(* IEC 61131-3 sources: RootPLC/conformance/cases/types, 56 files *)

(* ---- err_struct_recursive.st ---- *)
(* spec: [types.derived.struct]
   expect: error RP0107 *)
TYPE N : STRUCT child : N; END_STRUCT; END_TYPE

(* ---- err_subrange_bounds.st ---- *)
(* spec: [types.derived.subrange]
   expect: error RP0108 *)
TYPE Bad : INT (10..0); END_TYPE

(* ---- ok_call_through_reference.st ---- *)
(* spec: [types.reference.alias] [pous.call.callee]
   expect: warning RP0118
   run: PRG_Main cycles=2
   assert: c.n = 4 *)
FUNCTION_BLOCK FB_Count
VAR_OUTPUT
    n : INT;
END_VAR
n := n + 1;
END_FUNCTION_BLOCK

PROGRAM PRG_Main
VAR
    c : FB_Count;
    r : REFERENCE TO FB_Count;
END_VAR
r REF= c;
r();          (* calls c through the reference *)
c();
END_PROGRAM

(* ---- err_array_bound_not_constant.st ---- *)
(* spec: [variables.constant-names]
   expect: error RP0108 *)
PROGRAM PRG_Main
VAR
    n : INT := 4;
    buffer : ARRAY[0..n] OF INT;
END_VAR
END_PROGRAM

(* ---- err_array_bounds.st ---- *)
(* spec: [types.derived.array]
   expect: error RP0108 *)
PROGRAM PRG_Main
VAR
    a : ARRAY[5..1] OF INT;
END_VAR

END_PROGRAM

(* ---- err_array_const_index.st ---- *)
(* spec: [types.derived.array]
   expect: error RP0109 *)
PROGRAM PRG_Main
VAR
    a : ARRAY[0..2] OF INT;
END_VAR
a[3] := 1;
END_PROGRAM

(* ---- err_const_overflow.st ---- *)
(* spec: [types.int.overflow]
   expect: error RP0101 *)
PROGRAM PRG_Main
VAR
    x : LINT := 9223372036854775807 + 1;
END_VAR

END_PROGRAM

(* ---- err_dint_to_real.st ---- *)
(* spec: [types.conversion.implicit]
   expect: error RP0103 *)
PROGRAM PRG_Main
VAR
    r : REAL;
    d : DINT;
END_VAR
r := d;
END_PROGRAM

(* ---- err_div_const_zero.st ---- *)
(* spec: [types.int.division]
   expect: error RP0101 *)
PROGRAM PRG_Main
VAR
    x : INT;
END_VAR
x := 5 / 0;
END_PROGRAM

(* ---- err_enum_ambiguous.st ---- *)
(* spec: [types.derived.enum]
   expect: error RP0106 *)
TYPE Mode : (Off, Manual, Auto); END_TYPE

TYPE Valve : (Closed, Auto); END_TYPE

PROGRAM PRG_Main
VAR
    i : INT;
END_VAR
i := TO_INT(Auto);   (* no expected enumeration: Mode#Auto or Valve#Auto? *)
END_PROGRAM

(* ---- err_enum_strict_assign.st ---- *)
(* spec: [types.derived.enum.integer]
   expect: error RP0103 *)
{attribute 'qualified_only'}
{attribute 'strict'}
TYPE StrictMode : (Idle, Busy);
END_TYPE

PROGRAM PRG_Main
VAR
    s : StrictMode;
    i : INT := 1;
END_VAR
s := i;       (* an integer variable cannot be stored in a strict enumeration *)
i := s + 1;   (* no arithmetic on a strict enumeration *)
END_PROGRAM

(* ---- err_generic_decl.st ---- *)
(* spec: [types.generic]
   expect: error RP0104 *)
PROGRAM PRG_Main
VAR
    x : ANY_INT;
END_VAR

END_PROGRAM

(* ---- err_implicit_narrowing.st ---- *)
(* spec: [types.conversion.implicit]
   expect: error RP0103 *)
PROGRAM PRG_Main
VAR
    si : SINT;
    i : INT := 1;
END_VAR
si := i;
END_PROGRAM

(* ---- err_index_non_array.st ---- *)
(* spec: [types.derived.array]
   expect: error RP0103 *)
(* Only arrays (and, as vendor forms, strings and references) can be
   indexed. *)
PROGRAM PRG_Main
VAR
    x : INT;
    y : INT;
END_VAR
y := x[0];
END_PROGRAM

(* ---- err_int_to_bool.st ---- *)
(* spec: [types.conversion.implicit]
   expect: error RP0103 *)
PROGRAM PRG_Main
VAR
    b : BOOL;
    i : INT := 1;
END_VAR
b := i;
END_PROGRAM

(* ---- err_literal_range.st ---- *)
(* spec: [types.literal.range]
   expect: error RP0102 *)
PROGRAM PRG_Main
VAR
    x : SINT := 200;
END_VAR

END_PROGRAM

(* ---- err_string_len_zero.st ---- *)
(* spec: [types.derived.string]
   expect: error RP0108 *)
PROGRAM PRG_Main
VAR
    s : STRING[0];
END_VAR

END_PROGRAM

(* ---- err_struct_name_equivalence.st ---- *)
(* spec: [types.equivalence] [types.derived.struct]
   expect: error RP0103 *)
TYPE A : STRUCT v : INT; END_STRUCT; END_TYPE
TYPE B : STRUCT v : INT; END_STRUCT; END_TYPE

PROGRAM PRG_Main
VAR
    a : A;
    b : B;
END_VAR
a := b;
END_PROGRAM

(* ---- err_subrange_const.st ---- *)
(* spec: [types.derived.subrange]
   expect: error RP0105 *)
TYPE Percent : INT (0..100); END_TYPE

PROGRAM PRG_Main
VAR
    p : Percent := 150;
END_VAR

END_PROGRAM

(* ---- err_unknown_type.st ---- *)
(* spec: [types.derived.alias]
   expect: error RP0111 *)
PROGRAM PRG_Main
VAR
    x : NoSuchType;
END_VAR

END_PROGRAM

(* ---- ok_alias.st ---- *)
(* spec: [types.derived.alias] [types.equivalence]
   expect: ok
   run: PRG_Main cycles=1
   assert: i = 10
   assert: s = 11 *)
TYPE Speed : INT := 10; END_TYPE

PROGRAM PRG_Main
VAR
    s : Speed;
    i : INT;
END_VAR
i := s;
s := i + 1;
END_PROGRAM

(* ---- ok_array.st ---- *)
(* spec: [types.derived.array]
   expect: ok
   run: PRG_Main cycles=1
   assert: a[2] = 7
   assert: a[0] = 0
   assert: m[2, 2] = TRUE *)
PROGRAM PRG_Main
VAR
    a : ARRAY[0..2] OF INT;
    m : ARRAY[1..2, 1..2] OF BOOL;
END_VAR
a[2] := 7;
m[2, 2] := TRUE;
END_PROGRAM

(* ---- ok_conv_to_string.st ---- *)
(* spec: [types.conversion.explicit]
   expect: ok
   run: PRG_Main cycles=1
   assert: a = '42'
   assert: b = '255'
   assert: c = 'T#1s500ms'
   assert: d = 'A'
   assert: e = 'TRUE'
   assert: f = '-7' *)
PROGRAM PRG_Main
VAR
    a, b, c, d, e, f : STRING;
    ch : CHAR := CHAR#'A';
END_VAR
a := INT_TO_STRING(42);
b := WORD_TO_STRING(16#FF);
c := TIME_TO_STRING(T#1500MS);
d := CHAR_TO_STRING(ch);
e := BOOL_TO_STRING(TRUE);
f := DINT_TO_STRING(-7);
END_PROGRAM

(* ---- ok_datetime_to_string.st ---- *)
(* spec: [types.conversion.explicit]
   expect: ok
   run: PRG_Main cycles=1
   assert: sDt = 'DT#2017-04-04-12:42:42'
   assert: sD = 'D#1999-12-31'
   assert: sTod = 'TOD#08:05:03.25'
   assert: sB = 'TRUE'
   assert: sI = '-42' *)
PROGRAM PRG_Main
VAR
    sDt, sD, sTod, sB, sI : STRING;
END_VAR
sDt := DT_TO_STRING(DT#2017-04-04-12:42:42);
sD := DATE_TO_STRING(D#1999-12-31);
sTod := TOD_TO_STRING(TOD#08:05:03.25);
sB := BOOL_TO_STRING(TRUE);
sI := INT_TO_STRING(-42);
END_PROGRAM

(* ---- ok_default_init.st ---- *)
(* spec: [types.elementary] [types.default-init]
   expect: ok
   run: PRG_Main cycles=1
   assert: b = FALSE
   assert: i = 0
   assert: u = 0
   assert: r = 0.0
   assert: w = 0
   assert: t = T#0s
   assert: lt = LT#0s
   assert: d = D#1970-01-01
   assert: s = ''
   assert: ws = "" *)
PROGRAM PRG_Main
VAR
    b : BOOL;
    i : INT;
    u : ULINT;
    r : LREAL;
    w : WORD;
    t : TIME;
    lt : LTIME;
    d : DATE;
    s : STRING;
    ws : WSTRING;
END_VAR

END_PROGRAM

(* ---- ok_enum.st ---- *)
(* spec: [types.derived.enum]
   expect: ok
   run: PRG_Main cycles=1
   assert: first = Mode#Off
   assert: m = Mode#Auto
   assert: i = 2 *)
TYPE Mode : (Off, Manual, Auto); END_TYPE

PROGRAM PRG_Main
VAR
    m : Mode;
    first : Mode;
    i : INT;
END_VAR
first := m;
m := Manual;
m := Mode#Auto;
i := TO_INT(m);
END_PROGRAM

(* ---- ok_enum_value_by_context.st ---- *)
(* spec: [types.derived.enum]
   expect: ok
   run: PRG_Main cycles=1
   assert: n = 2
   assert: hit = TRUE
   assert: m = Motor#RUN
   assert: d = Door#OPEN *)
TYPE Motor : (IDLE, RUN, FAULT);
END_TYPE

TYPE Door : (IDLE, OPEN, CLOSED);
END_TYPE

FUNCTION F_Open : BOOL
VAR_INPUT
    d : Door;
END_VAR
F_Open := d = OPEN;
END_FUNCTION

PROGRAM PRG_Main
VAR
    m : Motor := IDLE;     (* initial value: Motor#IDLE *)
    d : Door;
    n : INT;
    hit : BOOL;
END_VAR
IF m = IDLE THEN           (* comparison: the other operand decides *)
    m := RUN;              (* assignment: the target decides *)
END_IF;
CASE m OF
    IDLE: n := 1;          (* CASE label: the selector decides *)
    RUN: n := 2;
END_CASE;
d := OPEN;
hit := F_Open(IDLE) = FALSE AND F_Open(d);   (* parameter decides *)
END_PROGRAM

(* ---- ok_explicit_conversion.st ---- *)
(* spec: [types.conversion.explicit]
   expect: ok
   run: PRG_Main cycles=1
   assert: a = 44
   assert: b = 3
   assert: c = -3
   assert: d = 127
   assert: e = -3 *)
PROGRAM PRG_Main
VAR
    a : SINT;
    b : INT;
    c : INT;
    d : SINT;
    e : INT;
END_VAR
a := INT_TO_SINT(300);
b := REAL_TO_INT(2.5);
c := REAL_TO_INT(-2.5);
d := LREAL_TO_SINT(1000.0);
e := TO_INT(SINT#-3);
END_PROGRAM

(* ---- ok_implicit_widening.st ---- *)
(* spec: [types.conversion.implicit]
   expect: ok
   run: PRG_Main cycles=1
   assert: i = -5
   assert: d = -5.0
   assert: w = 15 *)
PROGRAM PRG_Main
VAR
    s : SINT := -5;
    i : INT;
    d : LREAL;
    b : BYTE := 16#0F;
    w : WORD;
END_VAR
i := s;
d := i;
w := b;
END_PROGRAM

(* ---- ok_int_division.st ---- *)
(* spec: [types.int.division]
   expect: ok
   run: PRG_Main cycles=1
   assert: a = -3
   assert: b = -1
   assert: c = 1 *)
PROGRAM PRG_Main
VAR
    a : INT;
    b : INT;
    c : INT;
END_VAR
a := -7 / 2;
b := -7 MOD 2;
c := 7 MOD -2;
END_PROGRAM

(* ---- ok_int_wrap.st ---- *)
(* spec: [types.int.overflow]
   expect: ok
   run: PRG_Main cycles=1
   assert: x = -128
   assert: u = 255 *)
PROGRAM PRG_Main
VAR
    x : SINT := 127;
    u : USINT := 0;
END_VAR
x := x + 1;
u := u - 1;
END_PROGRAM

(* ---- ok_real_no_fault.st ---- *)
(* spec: [types.real]
   expect: ok
   run: PRG_Main cycles=1
   assert: big = TRUE *)
PROGRAM PRG_Main
VAR
    r : LREAL := 1.0;
    big : BOOL;
END_VAR
r := r / 0.0;
big := r > 1.0E308;
END_PROGRAM

(* ---- ok_reference.st ---- *)
(* spec: [types.reference]
   expect: ok
   run: PRG_Main cycles=1
   assert: x = 9 *)
PROGRAM PRG_Main
VAR
    x : INT := 5;
    r : REF_TO INT;
END_VAR
r := REF(x);
r^ := 9;
END_PROGRAM

(* ---- ok_string_truncate.st ---- *)
(* spec: [types.derived.string]
   expect: ok
   run: PRG_Main cycles=1
   assert: s = 'abcde' *)
PROGRAM PRG_Main
VAR
    s : STRING[5];
    t : STRING := 'abcdefgh';
END_VAR
s := t;
END_PROGRAM

(* ---- ok_struct.st ---- *)
(* spec: [types.derived.struct] [types.reference]
   expect: ok
   run: PRG_Main cycles=1
   assert: p.x = 1
   assert: p.y = 0
   assert: n.next = NULL *)
TYPE Point : STRUCT x : INT := 1; y : INT; END_STRUCT; END_TYPE
TYPE Node : STRUCT next : REF_TO Node; v : INT; END_STRUCT; END_TYPE

PROGRAM PRG_Main
VAR
    p : Point;
    n : Node;
END_VAR

END_PROGRAM

(* ---- ok_subrange.st ---- *)
(* spec: [types.derived.subrange]
   expect: ok
   run: PRG_Main cycles=1
   assert: first = 0
   assert: p = 50 *)
TYPE Percent : INT (0..100); END_TYPE

PROGRAM PRG_Main
VAR
    p : Percent;
    first : INT;
END_VAR
first := p;
p := 50;
END_PROGRAM

(* ---- ok_time_arithmetic.st ---- *)
(* spec: [types.time.arith]
   expect: ok
   run: PRG_Main cycles=1
   assert: t1 = TOD#08:30:00
   assert: t2 = TOD#23:30:00
   assert: d1 = DT#2026-11-04-12:01:30
   assert: d2 = DT#2026-11-04-11:59:00
   assert: dur1 = T#90000ms
   assert: dur2 = T#86400000ms
   assert: dur3 = T#3600000ms
   assert: lt = LTOD#00:00:01 *)
PROGRAM PRG_Main
VAR
    t1, t2 : TOD;
    d1, d2 : DT;
    dur1, dur2, dur3 : TIME;
    lt : LTOD;
END_VAR
t1 := TOD#08:00:00 + T#30M;
t2 := TOD#00:30:00 - T#1H;                        (* wraps around midnight *)
d1 := DT#2026-11-04-12:00:00 + T#1M30S500MS;      (* whole seconds *)
d2 := DT#2026-11-04-12:00:00 - T#1M;
dur1 := DT#2026-11-04-12:01:30 - DT#2026-11-04-12:00:00;
dur2 := D#2026-11-05 - D#2026-11-04;
dur3 := TOD#13:00:00 - TOD#12:00:00;
lt := LTOD#23:59:59 + LT#2S;
END_PROGRAM

(* ---- ok_time_conversions.st ---- *)
(* spec: [types.conversion.explicit] [types.conversion.implicit]
   expect: ok
   run: PRG_Main cycles=1
   assert: toL = LT#3ms
   assert: toT = T#1ms
   assert: viaTo = T#10ms
   assert: widened = LT#250ms
   assert: initL = LT#2s
   assert: atLdt = LDT#2026-01-01-10:00:00
   assert: atDt = DT#2026-01-01-10:00:00
   assert: atLtod = LTOD#12:30:00
   assert: gt = TRUE
   assert: eq = TRUE
   assert: later = TRUE
   assert: biggest = LT#2ms
   assert: ns = 1000000 *)
PROGRAM PRG_Main
VAR
    t : TIME := T#250ms;
    initL : LTIME := T#2s;
    toL, widened, biggest : LTIME;
    toT, viaTo : TIME;
    atLdt : LDT;
    atDt : DT;
    atLtod : LTOD;
    gt, eq, later : BOOL;
    ns : ULINT;
END_VAR
toL := TIME_TO_LTIME(T#3ms);
toT := LTIME_TO_TIME(LT#1500us);
viaTo := TO_TIME(TO_LTIME(UDINT#100000 * 100));
widened := t;
atLdt := DT#2026-01-01-10:00:00;
atDt := TO_DT(LDT#2026-01-01-10:00:00);
atLtod := TOD#12:30:00;
gt := T#2ms > LT#1ms;
eq := T#2ms = LT#2ms;
later := DT#2026-01-01-00:00:00 > LDT#2025-01-01-00:00:00;
biggest := MAX(T#2ms, LT#1ms);
ns := LTIME_TO_ULINT(T#1ms);
END_PROGRAM

(* ---- ok_to_string_forms.st ---- *)
(* spec: [types.conversion.explicit]
   expect: ok
   run: PRG_Main cycles=1
   assert: r1 = '0.1'
   assert: r2 = '-3.402823E38'
   assert: r3 = '1.0'
   assert: l1 = '123456789.0'
   assert: l2 = '1E-7'
   assert: t1 = 'T#49d17h2m47s295ms'
   assert: t2 = 'T#1s500ms'
   assert: t3 = 'T#0ms'
   assert: t4 = 'LT#1ms500us' *)
PROGRAM PRG_Main
VAR
    r1, r2, r3, l1, l2 : STRING;
    t1, t2, t3, t4 : STRING;
END_VAR
r1 := REAL_TO_STRING(REAL#0.1);
r2 := REAL_TO_STRING(REAL#-3.402823E38);
r3 := REAL_TO_STRING(REAL#1.0);
l1 := LREAL_TO_STRING(123456789.0);
l2 := LREAL_TO_STRING(1.0E-7);
t1 := TIME_TO_STRING(T#49d17h2m47s295ms);
t2 := TIME_TO_STRING(T#1500ms);
t3 := TIME_TO_STRING(T#0ms);
t4 := LTIME_TO_STRING(LTIME#1500us);
END_PROGRAM

(* ---- ok_untyped_literal.st ---- *)
(* spec: [types.literal.untyped]
   expect: ok
   run: PRG_Main cycles=1
   assert: u = 255
   assert: r = 3.0 *)
PROGRAM PRG_Main
VAR
    u : USINT := 255;
    r : REAL := 3;
END_VAR

END_PROGRAM

(* ---- warn_adr.st ---- *)
(* spec: [types.reference]
   expect: warning RP0117
   run: PRG_Main cycles=1
   assert: v = 9 *)
PROGRAM PRG_Main
VAR
    x : INT := 4;
    r : REF_TO INT;
    v : INT;
END_VAR
r := ADR(x);
r^ := 9;
v := x;
END_PROGRAM

(* ---- warn_array_bound_enum.st ---- *)
(* spec: [variables.constant-names] [scope.vendor-forms]
   expect: warning RP0135
   run: PRG_Main cycles=1
   assert: lo = 1
   assert: hi = 3
   assert: n = 3 *)
TYPE ST_Lanes :
STRUCT
    speed : ARRAY[E_Lane.Nr1..E_Lane.Nr3] OF INT;
END_STRUCT;
END_TYPE

TYPE E_Lane : (Nr1 := 1, Nr2, Nr3); END_TYPE

PROGRAM PRG_Main
VAR
    lanes : ARRAY[E_Lane.Nr1..E_Lane.Nr3] OF INT;
    lanes2 : ST_Lanes;
    lo, hi, n : DINT;
END_VAR
lo := LOWER_BOUND(lanes, 1);
hi := UPPER_BOUND(lanes, 1);
n := UPPER_BOUND(lanes2.speed, 1);
END_PROGRAM

(* ---- warn_enum_as_integer.st ---- *)
(* spec: [types.derived.enum.integer]
   expect: warning RP0129
   run: PRG_Main cycles=1
   assert: n = 2
   assert: plus = 3
   assert: next = Mode#Auto
   assert: same = TRUE
   assert: k = 1
   assert: fromInt = Mode#Manual
   assert: big = TRUE *)
TYPE Mode : (Off, Manual, Auto);
END_TYPE

TYPE Level : (Low, Mid, High);
END_TYPE

{attribute 'strict'}
TYPE StrictMode : (Idle, Busy);
END_TYPE

PROGRAM PRG_Main
VAR
    m : Mode := Mode#Auto;
    n : INT;
    plus : INT;
    next : Mode;
    same : BOOL;
    k : INT;
    fromInt : Mode;
    i : INT := 1;
    s : StrictMode;
    big : BOOL;
END_VAR
n := m;                           (* value as integer *)
plus := Mode#Auto + 1;            (* arithmetic on a non-strict enumeration *)
next := Mode#Manual + 1;          (* integer stored in a non-strict enumeration *)
same := Mode#Auto = Level#High;   (* compared as integers *)
s := StrictMode#Busy;
k := s;                           (* a strict value still reads as an integer *)
big := s > 0;
fromInt := i;
END_PROGRAM

(* ---- warn_enum_base_type_after.st ---- *)
(* spec: [types.derived.enum]
   expect: warning RP0115
   run: PRG_Main cycles=1
   assert: n = 10 *)
TYPE E_Mode : (Off := 0, Manual := 5, Auto := 10) UINT; END_TYPE

PROGRAM PRG_Main
VAR
    m : E_Mode := E_Mode#Auto;
    n : INT;
END_VAR
n := TO_INT(m);
END_PROGRAM

(* ---- warn_enum_dot_value.st ---- *)
(* spec: [types.derived.enum]
   expect: warning RP0122
   run: PRG_Main cycles=1
   assert: n = 10
   assert: same = TRUE
   assert: k = 1 *)
TYPE E_Mode : (Off := 0, Manual := 5, Auto := 10); END_TYPE

NAMESPACE Plant
TYPE E_Valve : (Closed, Open); END_TYPE
END_NAMESPACE

PROGRAM PRG_Main
VAR
    m : E_Mode := E_Mode.Auto;
    v : Plant.E_Valve;
    n, k : INT;
    same : BOOL;
END_VAR
n := TO_INT(m);
same := m = E_Mode#Auto;
v := Plant.E_Valve.Open;
k := TO_INT(v);
END_PROGRAM

(* ---- warn_enum_to_int.st ---- *)
(* spec: [types.derived.enum] [types.derived.enum.integer]
   expect: warning RP0129
   run: PRG_Main cycles=1
   assert: i = 2
   assert: j = 2 *)
TYPE Mode : (Off, Manual, Auto); END_TYPE

PROGRAM PRG_Main
VAR
    m : Mode := Mode#Auto;
    i, j : INT;
END_VAR
i := m;          (* accepted with RP0129 (CODESYS / TwinCAT) *)
j := TO_INT(m);  (* the portable spelling *)
END_PROGRAM

(* ---- warn_index_string_and_pointer.st ---- *)
(* spec: [types.derived.array] [types.reference] [scope.vendor-forms]
   expect: warning RP0135
   run: PRG_Main cycles=1
   assert: third = 40
   assert: changed = 99
   assert: first = 97
   assert: past = 0
   assert: text = 'aBcd'
   assert: cut = 'a'
   assert: wide = 121 *)
(* CODESYS / TwinCAT character access s[i] and pointer index p[i]. *)
PROGRAM PRG_Main
VAR
    a       : ARRAY[0..3] OF INT := [10, 20, 30, 40];
    r       : REF_TO INT;
    s       : STRING[5] := 'abc';
    w       : WSTRING[4] := "xy";
    third   : INT;
    changed : INT;
    first   : BYTE;
    past    : BYTE;
    text    : STRING[5];
    cut     : STRING[5];
    wide    : WORD;
END_VAR
r := REF(a[1]);
third := r[2];
r[1] := 99;
changed := a[2];
first := s[0];
past := s[3];
s[1] := 66;
s[3] := 100;
text := s;
s[1] := 0;
cut := s;
wide := w[1];
END_PROGRAM

(* ---- warn_pointer_to.st ---- *)
(* spec: [types.reference]
   expect: warning RP0116
   run: PRG_Main cycles=1
   assert: v = 7 *)
PROGRAM PRG_Main
VAR
    x : INT := 7;
    p : POINTER TO INT;
    v : INT;
END_VAR
p := REF(x);
v := p^;
END_PROGRAM

(* ---- warn_reference_alias.st ---- *)
(* spec: [types.reference.alias]
   expect: warning RP0118 RP0006
   run: PRG_Main cycles=1
   assert: x = 12
   assert: v = 12
   assert: valid
   assert: NOT before *)
PROGRAM PRG_Main
VAR
    x : INT := 2;
    r : REFERENCE TO INT;
    v : INT;
    valid, before : BOOL;
END_VAR
before := __ISVALIDREF(r);
r REF= x;
valid := __ISVALIDREF(r);
r := r + 10;
v := r;
END_PROGRAM

(* ---- warn_same_size_bits.st ---- *)
(* spec: [types.conversion.vendor]
   expect: warning RP0126
   run: PRG_Main cycles=1
   assert: x = 3
   assert: y = 6 *)
PROGRAM PRG_Main
VAR
    w : DWORD := 5;
    u : UDINT := 3;
    x, y : DWORD;
END_VAR
x := u;
y := w XOR u;
END_PROGRAM

(* ---- warn_string_length_parens.st ---- *)
(* spec: [types.derived.string]
   expect: warning RP0112
   run: PRG_Main cycles=1
   assert: n = 3 *)
PROGRAM PRG_Main
VAR
    s : STRING(3) := 'abc';
    w : WSTRING(10);
    t : STRING := 'abcdef';
    n : INT;
END_VAR
s := t;
n := LEN(s);
END_PROGRAM

(* ---- warn_string_too_long.st ---- *)
(* spec: [types.derived.string]
   expect: warning RP0110 *)
PROGRAM PRG_Main
VAR
    s : STRING[3] := 'abcdef';
END_VAR

END_PROGRAM

(* ---- warn_struct_empty.st ---- *)
(* spec: [types.derived.struct] [scope.vendor-forms]
   expect: warning RP0134 *)
TYPE ST_Placeholder :
STRUCT
END_STRUCT;
END_TYPE

PROGRAM PRG_Main
VAR
    s : ST_Placeholder;
END_VAR
END_PROGRAM

(* ---- warn_struct_extends.st ---- *)
(* spec: [types.derived.struct] [scope.vendor-forms]
   expect: warning RP0134
   run: PRG_Main cycles=1
   assert: a = 5
   assert: b = 2 *)
TYPE
    ST_Base : STRUCT
        id : INT := 5;
    END_STRUCT;
    ST_Item EXTENDS ST_Base : STRUCT
        qty : INT := 2;
    END_STRUCT;
END_TYPE

PROGRAM PRG_Main
VAR
    it : ST_Item;
    a, b : INT;
END_VAR
a := it.id;
b := it.qty;
END_PROGRAM

(* ---- warn_union.st ---- *)
(* spec: [types.derived.union] [scope.vendor-forms]
   libraries: TwinCAT_BuiltIns
   expect: warning RP0134
   run: PRG_Main cycles=1
   assert: n = 8 *)
TYPE U_Value :
UNION
    asReal : LREAL;
    asBits : LWORD;
    asBytes : ARRAY[0..3] OF BYTE;
END_UNION;
END_TYPE

PROGRAM PRG_Main
VAR
    u : U_Value;
    n : UDINT;
END_VAR
n := SIZEOF(u);
END_PROGRAM

(* ---- warn_vendor_conversions.st ---- *)
(* spec: [types.conversion.vendor]
   expect: warning RP0126 RP0127
   run: PRG_Main cycles=1
   assert: w = 0
   assert: m = 4
   assert: v = 4
   assert: flag = FALSE
   assert: isNull = TRUE *)
PROGRAM PRG_Main
VAR
    w : DWORD := 16#FFFFFFFF;
    u : UDINT := 12;
    m : UDINT;
    i : BYTE := 3;
    arr : ARRAY[0..3] OF INT := [1, 2, 3, 4];
    v : INT;
    flag : BOOL := 1;
    p : REF_TO INT := 0;
    isNull : BOOL;
END_VAR
w := w + 1;
m := u AND 4;
v := arr[i];
flag := 0;
isNull := p = NULL;
END_PROGRAM
